FUNCTION_BLOCK FB_GFX4IR_REF
VAR_INPUT
	Gfx4IRToPlc			AT %I*:ARRAY[1..4] OF ST_GFX4IRTOPLC;
END_VAR
VAR_OUTPUT
	PlcToGfx4IR			AT %Q*:ARRAY[1..4] OF ST_PLCTOGFX4IR;
END_VAR
VAR
END_VAR

;

END_FUNCTION_BLOCK

(* stored: Version 1.1.0.1, ProductVersion 3.1.4024.15
   POU FB_GFX4IR_REF: Id {3a65c466-5440-42ff-82af-e32ee13b9ba8}, SpecialFunc None *)
